// TIA Portal V20 export
DATA_BLOCK "T7_Std"   // DB44902
{ S7_Optimized_Access := 'FALSE' }
AUTHOR : IA
FAMILY : PRUEBA
VERSION : 0.1
// Tanda 3: DB de acceso estándar para PEEK/POKE (número fijo 44902)
// stored: AutoNumber false
   VAR
      W : Word;   // Destino de POKE (byte 0)
      Relleno : Array[0..9] of Byte;
   END_VAR
BEGIN
END_DATA_BLOCK
